// TIA Portal V21 export
// export: Created 2026-10-14T03:09:01.8081687Z, ExportSetting WithDefaults, DisplayName Totally Integrated Automation Portal, DisplayVersion V21, DisplayName STEP 7 Professional, DisplayVersion V21, DisplayName STEP 7 Safety, DisplayVersion V21, DisplayName Tech WebApplication, DisplayVersion V21, DisplayName WinCC Basic/Comfort/Advanced, DisplayVersion V21, DisplayName WinCC Unified, DisplayVersion V21
TagTable "Template"
  MainNavigationState : Int  (1 s, start 1)
  SubNavigationState : Int  (1 s, start 1)
  CurrentUserName : WString  (1 s)
  DiagState : Int  (1 s)
  PopUpBackground : Bool  (1 s)
  UserName : WString  (1 s)
  Password : WString  (1 s)
  UserIsLoggedIn : Bool  (1 s)
  CodeView : Bool  (1 s)
  Brightness : Int  (1 s, start 100)
  CurrentLanguage : Bool  (1 s)
  CurrentRecipeName : WString  (1 s)
  CurrentMachineState : Int  (1 s)
  OptionPanelNavigationState : Int  (1 s, start 1)
  ButtonDown : Bool  (1 s)
  ThirdLevelNavigationState : Int  (1 s, start 1)
  StartScreenName : WString  (1 s)
  InScreenTabState : Int  (1 s, start 0)
  DummyTagBool : Bool  (1 s)
  DummyTagInt1 : Int  (1 s)
  DummyTagInt2 : Int  (1 s)
  DummyTagInt3 : Int  (1 s)
  DummyDeltaReal : LReal  (1 s, start 0.1)
  DummTagReal1 : LReal  (1 s)
  DummyDeltaInt : Int  (1 s, start 1)
